SUBAPPLICATION E_PERMIT_INVERT_2 (* 2-Kanal invertiertes Event-Freigabe-Gate (je Kanal F_NOT_BOOL_INIT + E_PERMIT) *)
  (* Standard: 61499-2; Description: Copyright (c) 2026 Meisterschulen am Ostbahnhof This program and the accompanying materials are made available under the terms of the Eclipse Public License 2.0 which is available at https://www.eclipse.org/legal/epl-2.0/ SPDX-License-Identifier: EPL-2.0 *)
  (* Version 1.1, 2026-11-11, Franz Höpfinger, Meisterschulen am Ostbahnhof, Je Kanal ein F_NOT_BOOL_INIT und ein E_PERMIT statt E_MUX/E_DEMUX mit gemeinsamem K: kamen zwei Kanaele in derselben Ereigniskette (z. B. E_SPLIT), ueberschrieb E_MUX das K, bevor E_DEMUX es las, und das erste Ereignis landete auf dem falschen Ausgang. *)
  (* Version 1.0, 2026-09-10, Franz Höpfinger, Meisterschulen am Ostbahnhof, initial implementation *)
  PACKAGE MyLib::sys;
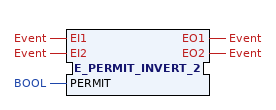
  EVENT_INPUT
    EI1; (* Event input channel 1 *)
    EI2; (* Event input channel 2 *)
  END_EVENT
  EVENT_OUTPUT
    EO1; (* Event output channel 1 *)
    EO2; (* Event output channel 2 *)
  END_EVENT
  VAR_INPUT
    PERMIT : BOOL; (* Invertierte Freigabebedingung *)
  END_VAR
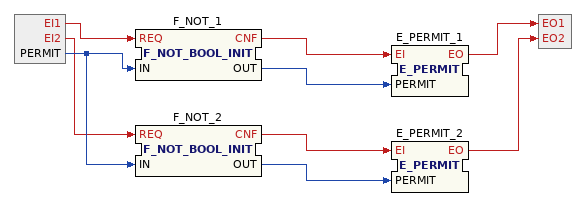
  FBS
    F_NOT_1 : iec61131::booleanOperators::F_NOT_BOOL_INIT;
    E_PERMIT_1 : iec61499::events::E_PERMIT;
    F_NOT_2 : iec61131::booleanOperators::F_NOT_BOOL_INIT;
    E_PERMIT_2 : iec61499::events::E_PERMIT;
  END_FBS
  EVENT_CONNECTIONS
    EI1 TO F_NOT_1.REQ;
    F_NOT_1.CNF TO E_PERMIT_1.EI;
    E_PERMIT_1.EO TO EO1;
    EI2 TO F_NOT_2.REQ;
    F_NOT_2.CNF TO E_PERMIT_2.EI;
    E_PERMIT_2.EO TO EO2;
  END_CONNECTIONS
  DATA_CONNECTIONS
    PERMIT TO F_NOT_1.IN;
    F_NOT_1.OUT TO E_PERMIT_1.PERMIT;
    PERMIT TO F_NOT_2.IN;
    F_NOT_2.OUT TO E_PERMIT_2.PERMIT;
  END_CONNECTIONS
END_SUBAPPLICATION
